(* IEC 61131-3 sources: plc-repo-template/tests/POUs/FB_F_Clamp_Test, 8 files *)

(* ---- FB_F_Clamp_Test.decl.st ---- *)
// Назначение: набор тестов CfUnit (coUnit 1.2.0.0) для F_Clamp — значение внутри
//             диапазона, ниже, выше, на границах, вырожденный диапазон и границы
//             в обратном порядке. Экземпляр объявлен в PRG_Tests: объявление
//             регистрирует набор в coUnit, вызывать его вручную не нужно.
// Автор:      kr0nsch
// Версия:     0.1.0
// Документ:   docs/TEST_REPORT.md
FUNCTION_BLOCK FB_F_Clamp_Test EXTENDS coUnit.FB_TestSuite
VAR CONSTANT
    // Ожидаемые значения не равны нулю: функция без реализации вернула бы 0,
    // и тест с ожиданием 0 прошёл бы ложно.
    R_LOW : REAL := 2.0;        // нижняя граница тестового диапазона
    R_HIGH : REAL := 10.0;      // верхняя граница тестового диапазона
    R_INSIDE : REAL := 5.0;     // значение внутри диапазона
    R_BELOW : REAL := -3.0;     // значение ниже диапазона
    R_ABOVE : REAL := 12.5;     // значение выше диапазона
    // F_Clamp возвращает один из своих аргументов без арифметики — сравнение точное
    R_DELTA : REAL := 0.0;
END_VAR

(* ---- AboveHighReturnsHigh.method.decl.st ---- *)
// Значение выше диапазона заменяется верхней границей.
METHOD PRIVATE AboveHighReturnsHigh
VAR
    rResult : REAL;     // результат F_Clamp
END_VAR

(* ---- AtHighBoundaryReturnsHigh.method.decl.st ---- *)
// Значение, равное верхней границе, возвращается без изменений.
METHOD PRIVATE AtHighBoundaryReturnsHigh
VAR
    rResult : REAL;     // результат F_Clamp
END_VAR

(* ---- AtLowBoundaryReturnsLow.method.decl.st ---- *)
// Значение, равное нижней границе, возвращается без изменений.
METHOD PRIVATE AtLowBoundaryReturnsLow
VAR
    rResult : REAL;     // результат F_Clamp
END_VAR

(* ---- BelowLowReturnsLow.method.decl.st ---- *)
// Значение ниже диапазона заменяется нижней границей.
METHOD PRIVATE BelowLowReturnsLow
VAR
    rResult : REAL;     // результат F_Clamp
END_VAR

(* ---- EqualBoundsReturnsBound.method.decl.st ---- *)
// Вырожденный диапазон (rLow = rHigh): результат всегда равен границе.
METHOD PRIVATE EqualBoundsReturnsBound
VAR
    rResult : REAL;     // результат F_Clamp
END_VAR

(* ---- InsideRangeReturnsValue.method.decl.st ---- *)
// Значение внутри диапазона возвращается без изменений.
METHOD PRIVATE InsideRangeReturnsValue
VAR
    rResult : REAL;     // результат F_Clamp
END_VAR

(* ---- LowGreaterThanHighSwapsBounds.method.decl.st ---- *)
// Границы в обратном порядке (rLow > rHigh) меняются местами — см. docs/ASSUMPTIONS.md.
METHOD PRIVATE LowGreaterThanHighSwapsBounds
VAR
    rResult : REAL;     // результат F_Clamp
END_VAR
